{attribute 'qualified_only'}
{attribute 'to_string'}
TYPE E_Anybus_RecipeType :
(
	eNone			:= 0,	// not selected
	eFlushOnly				:= 1,	// CIP1
	eDetergent				:= 2,	// CIP1, CIP2, CIP3
	eDetergentOnly			:= 3,	// CIP2, CIP3
	eDisinfectionOnly		:= 4,	// CIP4, CIP5
	eDetergentDisinfection	:= 5,	// CIP2 .. CIP5
	eFull					:= 6	// CIP1 .. CIP5, codes proposed to GAD 02.11.2026
);
END_TYPE

(* stored: Version 1.1.0.1, ProductVersion 3.1.4026.20
   DUT E_Anybus_RecipeType: Id {2496285c-e348-414b-9c1d-31a8acdde51c} *)
